Staubli VAL3: bIsHome.pgx

program bIsHome(jointRx x_jHome, bool& x_bAtHome)
begin
  //判断当前位置是否为Home点
  x_bAtHome=(abs((herej()-x_jHome))<{4,4,4,4,4,4})
end
